// TIA Portal V20 export
// export: Created 2026-10-12T05:26:51.415726Z, ExportSetting WithDefaults, DisplayName Totally Integrated Automation Portal, DisplayVersion V20, DisplayName TIA Portal Openness, DisplayVersion V20, DisplayName TIA Portal Teamcenter Gateway, DisplayVersion V20, DisplayName TIA Portal Version Control Interface, DisplayVersion V20, DisplayName SINAMICS Startdrive Advanced, DisplayVersion V20 SP1 Update 2, DisplayName SINAMICS Startdrive G110M, G120, G120C, G120D, G120P, G115D, DisplayVersion V20 SP1 Update 2, DisplayName SINAMICS Startdrive G130, G150, S120, S150, SINAMICS MV, G220, S200, S210, DisplayVersion V20 SP1 Update 2, DisplayName STEP 7 Professional, DisplayVersion V20, DisplayName STEP 7 Safety, DisplayVersion V20, DisplayName WinCC Basic/Comfort/Advanced, DisplayVersion V20, DisplayName WinCC Professional, DisplayVersion V20, DisplayName WinCC Unified, DisplayVersion V20
FUNCTION "FRK_ManualCommon" : Void   // FC81, SCL
{ S7_Optimized_Access := 'TRUE' }
VERSION : 0.1
// stored: AutoNumber true, IsIECCheckEnabled false, SetENOAutomatically false, UDAEnableTagReadback false
   VAR_INPUT
      Core : "FRK_Core";
      Unit : "FRK_Unit";
      Status : "ST_ModuleStatus";
   END_VAR
   VAR_IN_OUT
      Report : "ST_ReleaseReport";
   END_VAR
BEGIN

   IF #Unit.Mode <> 1 OR #Unit.ModePending THEN
       "FRK_ReleaseReason"(Report := #Report,
                           Description := WSTRING#'std.release.manualModeRequired',
                           Reason := 2002,
                           Path := STRING_TO_WSTRING(#Status.Name),
                           Kind := 0);
   END_IF;
   IF #Core.Exec <> 0 OR #Unit.Clearing OR #Unit.FaultLatched THEN
       "FRK_ReleaseReason"(Report := #Report,
                           Description := WSTRING#'std.error.hmiRequestRejected',
                           Reason := 2011,
                           Path := STRING_TO_WSTRING(#Status.Name),
                           Kind := 4);
   END_IF;
   IF #Unit.AlarmBlocking THEN
       "FRK_ReleaseReason"(Report := #Report,
                           Description := WSTRING#'std.release.manualReset',
                           Reason := 0,
                           Path := STRING_TO_WSTRING(#Status.Name),
                           Kind := 2);
   END_IF;
   IF NOT #Unit.Permit THEN
       "FRK_ReleaseReason"(Report := #Report,
                           Description := #Unit.PermitDiag.Description,
                           Reason := #Unit.PermitDiag.ReasonCode,
                           Path := #Unit.PermitDiag.SourcePath,
                           Kind := 3);
   END_IF;
END_FUNCTION
